(*
SPDX-FileCopyrightText: © 2026 Oleksandr Tiutyk <trofimich@gmail.com>
SPDX-License-Identifier: MIT
License: https://opensource.org/license/mit
*)

(*!
<summary>Beckhoff EL3413/EL3433 auxiliary measurement selectors.</summary>
<description>
Represents RxPDO 0x1603: Index at 0x7030:01 and Channel at 0x7030:02, both UINT8.
Select a combination supported by the device/firmware. Selection takes effect asynchronously;
wait for both acknowledged input selectors and valid input status before interpreting auxiliary Value.
Link fields individually and use one owner task for writes; externally synchronize other access.
When used for I/O, link located fields or their containing buffers to the matching selected PDOs.
The record is not a packed wire buffer; compiler padding is not part of the device specification.
Unlinked/default values do not prove valid I/O. The caller evaluates bus/channel validity before use.
Use one owner task per instance and externally synchronize other access; multi-field snapshots are not atomic.
Copies store data without creating hardware links. Keep borrowed field references valid while consumers are bound.
This passive record performs no validation, synchronization, configuration or protocol advancement.
</description>
*)
TYPE POWER_MEASUREMENT_AUXILIARY_OUTPUT_CHANNEL :
STRUCT
	Index AT %Q* : USINT;
	Channel AT %Q* : USINT;
END_STRUCT
END_TYPE

(* stored: Version 1.1.0.1
   DUT POWER_MEASUREMENT_AUXILIARY_OUTPUT_CHANNEL: Id {c8ba096f-ece7-433b-9679-aa57ac825437} *)
